(* IEC 61131-3 sources: rusty/compiler/plc_cfc/fixtures/blocks/invalid/function_inout_negated, 1 file *)

(* ---- addInto.st ---- *)
FUNCTION addInto : DINT
VAR_INPUT
    delta : DINT;
END_VAR
VAR_IN_OUT
    acc : DINT;
END_VAR
    acc := acc + delta;
    addInto := acc;
END_FUNCTION
